// TIA Portal V19 export
FUNCTION_BLOCK "MOTOR_FB1"   // FB6, LAD
{ S7_Optimized_Access := 'FALSE' }
// stored: SetENOAutomatically false
   VAR_INPUT
      TRIP : Bool;
   END_VAR
   VAR_OUTPUT
      OP_FBK_ERROR : Bool;
      CL_FBK_ERROR : Bool;
      AUTO_MODE : Bool;
      MANUAL_MODE : Bool;
      SEMI_AUTO_MODE : Bool;
      "START/STOPCMD" : Bool;
      STATUS : Int;
   END_VAR
   VAR_IN_OUT
      "MANUAL SELECTION" : Bool;
      SEMI : Bool;
      "MANUAL START" : Bool;
      "AUTO START" : Bool;
      "FEEDBACK RUN" : Bool;
      TRIPPED : Bool;
      REMOTE : Bool;
      RESET : Bool;
      INTERLOCK : Bool;
      "WAITING TIME" : DInt;
   END_VAR
   VAR
      "TIMER" { S7_SetPoint := 'True'} : IEC_TIMER;
      MON_ERROR : Bool;
      INTERLOCK_ACTIVE : Bool;
   END_VAR
   // "TIMER".PT := T#10S;
   VAR_TEMP   // added for the SCL form of the ladder/FBD networks
      _w1 : Bool;
   END_VAR
BEGIN

REGION Network 1: MODE SELECTION
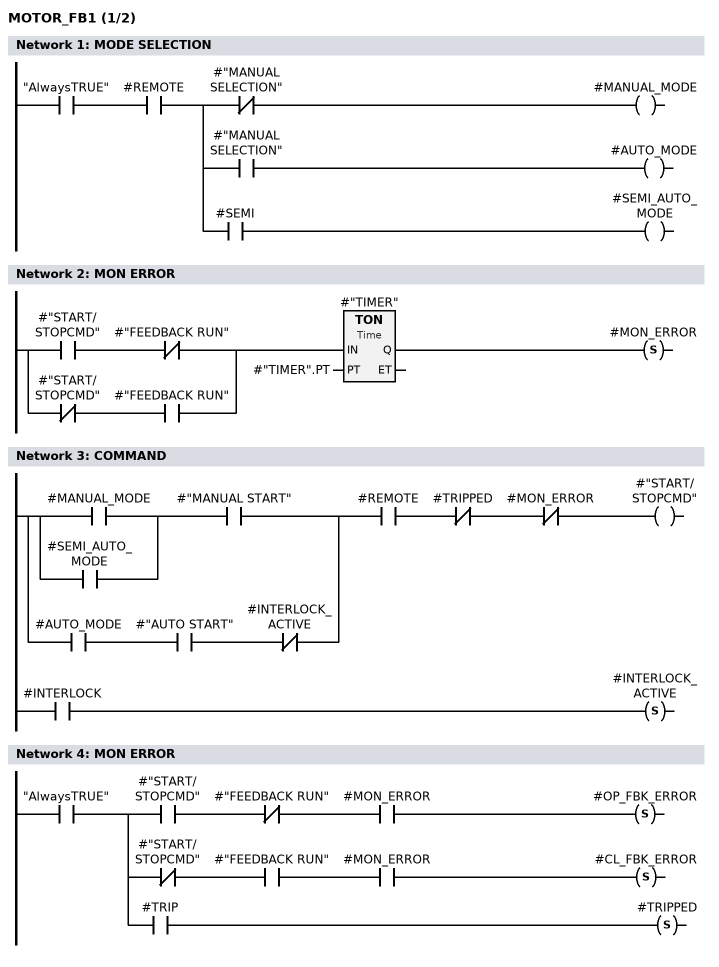
   RUNG wire#powerrail
      Contact( "AlwaysTRUE" )
      Contact( #REMOTE )
      wire#w1
      I_Contact( #"MANUAL SELECTION" )
      Coil( #MANUAL_MODE )
   END_RUNG
   RUNG wire#w1
      Contact( #"MANUAL SELECTION" )
      Coil( #AUTO_MODE )
   END_RUNG
   RUNG wire#w1
      Contact( #SEMI )
      Coil( #SEMI_AUTO_MODE )
   END_RUNG
   // the same network as SCL:
   #_w1 := "AlwaysTRUE" AND #REMOTE;
   #MANUAL_MODE := #_w1 AND NOT #"MANUAL SELECTION";
   #AUTO_MODE := #_w1 AND #"MANUAL SELECTION";
   #SEMI_AUTO_MODE := #_w1 AND #SEMI;
END_REGION

REGION Network 2: MON ERROR
   RUNG wire#powerrail
      Contact( #"START/STOPCMD" )
      I_Contact( #"FEEDBACK RUN" )
      wire#w1
      { S7_Templates := "time_type := Time" } #"TIMER".TON(pt := #"TIMER".PT, et =>)
      S_Coil( #MON_ERROR )
   END_RUNG
   RUNG wire#powerrail
      I_Contact( #"START/STOPCMD" )
      Contact( #"FEEDBACK RUN" )
   END_RUNG wire#w1
   // the same network as SCL:
   #"TIMER".TON(IN := (#"START/STOPCMD" AND NOT #"FEEDBACK RUN") OR (NOT #"START/STOPCMD" AND #"FEEDBACK RUN"),
                PT := #"TIMER".PT);
   IF #"TIMER".Q THEN #MON_ERROR := TRUE; END_IF;
END_REGION

REGION Network 3: COMMAND
   RUNG wire#powerrail
      Contact( #MANUAL_MODE )
      wire#w1
      Contact( #"MANUAL START" )
      wire#w2
      Contact( #REMOTE )
      I_Contact( #TRIPPED )
      I_Contact( #MON_ERROR )
      Coil( #"START/STOPCMD" )
   END_RUNG
   RUNG wire#powerrail
      Contact( #SEMI_AUTO_MODE )
   END_RUNG wire#w1
   RUNG wire#powerrail
      Contact( #AUTO_MODE )
      Contact( #"AUTO START" )
      I_Contact( #INTERLOCK_ACTIVE )
   END_RUNG wire#w2
   RUNG wire#powerrail
      Contact( #INTERLOCK )
      S_Coil( #INTERLOCK_ACTIVE )
   END_RUNG
   // the same network as SCL:
   #"START/STOPCMD" := (((#MANUAL_MODE OR #SEMI_AUTO_MODE) AND #"MANUAL START") OR (#AUTO_MODE AND #"AUTO START" AND NOT #INTERLOCK_ACTIVE)) AND #REMOTE AND NOT #TRIPPED AND NOT #MON_ERROR;
   IF #INTERLOCK THEN #INTERLOCK_ACTIVE := TRUE; END_IF;
END_REGION

REGION Network 4: MON ERROR
   RUNG wire#powerrail
      Contact( "AlwaysTRUE" )
      wire#w1
      Contact( #"START/STOPCMD" )
      I_Contact( #"FEEDBACK RUN" )
      Contact( #MON_ERROR )
      S_Coil( #OP_FBK_ERROR )
   END_RUNG
   RUNG wire#w1
      I_Contact( #"START/STOPCMD" )
      Contact( #"FEEDBACK RUN" )
      Contact( #MON_ERROR )
      S_Coil( #CL_FBK_ERROR )
   END_RUNG
   RUNG wire#w1
      Contact( #TRIP )
      S_Coil( #TRIPPED )
   END_RUNG
   // the same network as SCL:
   IF "AlwaysTRUE" AND #"START/STOPCMD" AND NOT #"FEEDBACK RUN" AND #MON_ERROR THEN
       #OP_FBK_ERROR := TRUE;
   END_IF;
   IF "AlwaysTRUE" AND NOT #"START/STOPCMD" AND #"FEEDBACK RUN" AND #MON_ERROR THEN
       #CL_FBK_ERROR := TRUE;
   END_IF;
   IF "AlwaysTRUE" AND #TRIP THEN #TRIPPED := TRUE; END_IF;
END_REGION

REGION Network 5: STATUS
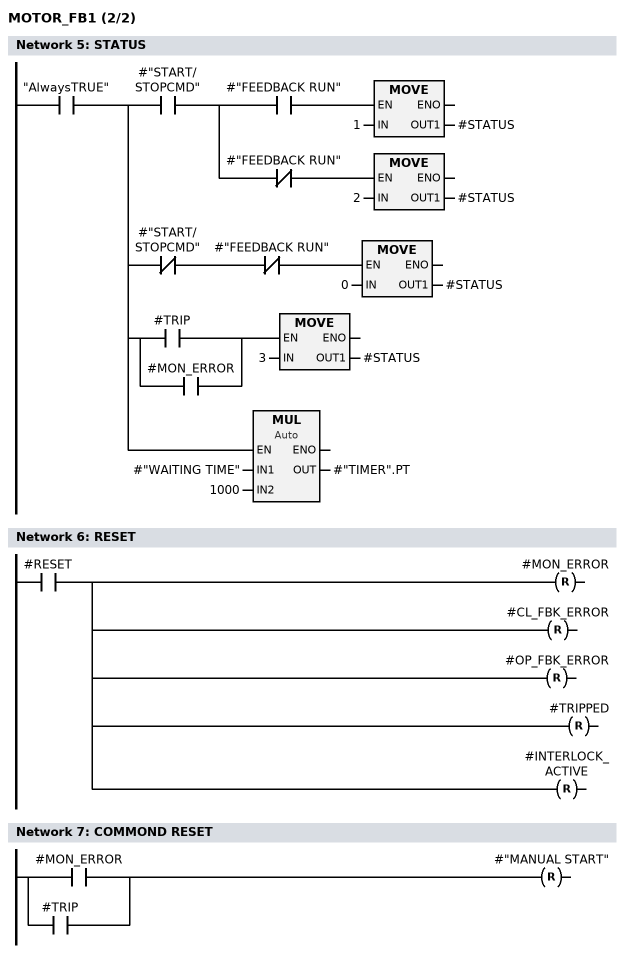
   RUNG wire#powerrail
      Contact( "AlwaysTRUE" )
      wire#w1
      Contact( #"START/STOPCMD" )
      wire#w2
      Contact( #"FEEDBACK RUN" )
      Move(in := 1, out1 => #STATUS)
   END_RUNG
   RUNG wire#w2
      I_Contact( #"FEEDBACK RUN" )
      Move(in := 2, out1 => #STATUS)
   END_RUNG
   RUNG wire#w1
      I_Contact( #"START/STOPCMD" )
      I_Contact( #"FEEDBACK RUN" )
      Move(in := 0, out1 => #STATUS)
   END_RUNG
   RUNG wire#w1
      Contact( #TRIP )
      wire#w3
      Move(in := 3, out1 => #STATUS)
   END_RUNG
   RUNG wire#w1
      Contact( #MON_ERROR )
   END_RUNG wire#w3
   RUNG wire#w1
      Mul(in1 := #"WAITING TIME", in2 := 1000, out => #"TIMER".PT)
   END_RUNG
   // the same network as SCL:
   #_w1 := "AlwaysTRUE" AND #"START/STOPCMD";
   IF #_w1 AND #"FEEDBACK RUN" THEN #STATUS := 1; END_IF;
   IF #_w1 AND NOT #"FEEDBACK RUN" THEN #STATUS := 2; END_IF;
   IF "AlwaysTRUE" AND NOT #"START/STOPCMD" AND NOT #"FEEDBACK RUN" THEN #STATUS := 0; END_IF;
   IF "AlwaysTRUE" AND (#TRIP OR #MON_ERROR) THEN #STATUS := 3; END_IF;
   IF "AlwaysTRUE" THEN #"TIMER".PT := #"WAITING TIME" * 1000; END_IF;
END_REGION

REGION Network 6: RESET
   RUNG wire#powerrail
      Contact( #RESET )
      wire#w1
      R_Coil( #MON_ERROR )
   END_RUNG
   RUNG wire#w1
      R_Coil( #CL_FBK_ERROR )
   END_RUNG
   RUNG wire#w1
      R_Coil( #OP_FBK_ERROR )
   END_RUNG
   RUNG wire#w1
      R_Coil( #TRIPPED )
   END_RUNG
   RUNG wire#w1
      R_Coil( #INTERLOCK_ACTIVE )
   END_RUNG
   // the same network as SCL:
   IF #RESET THEN
       #MON_ERROR := FALSE;
       #CL_FBK_ERROR := FALSE;
       #OP_FBK_ERROR := FALSE;
       #TRIPPED := FALSE;
       #INTERLOCK_ACTIVE := FALSE;
   END_IF;
END_REGION

REGION Network 7: COMMOND RESET
   RUNG wire#powerrail
      Contact( #MON_ERROR )
      wire#w1
      R_Coil( #"MANUAL START" )
   END_RUNG
   RUNG wire#powerrail
      Contact( #TRIP )
   END_RUNG wire#w1
   // the same network as SCL:
   IF #MON_ERROR OR #TRIP THEN #"MANUAL START" := FALSE; END_IF;
END_REGION
END_FUNCTION_BLOCK
